FUNCTION_BLOCK IMU_STREAM
  {SET_ATTRIBUTE(OpcUa, SERVICE)}
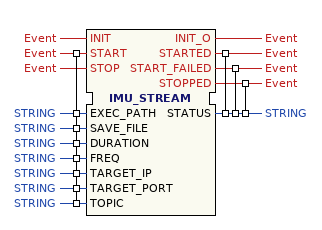
  EVENT_INPUT
    INIT;
    START WITH EXEC_PATH, SAVE_FILE, DURATION, FREQ, TARGET_IP, TARGET_PORT, TOPIC;
    STOP;
  END_EVENT
  EVENT_OUTPUT
    INIT_O;
    STARTED WITH STATUS;
    START_FAILED WITH STATUS;
    STOPPED WITH STATUS;
  END_EVENT
  VAR_INPUT
    EXEC_PATH : STRING; {SET_ATTRIBUTE(OpcUa, Variable)}
    SAVE_FILE : STRING; {SET_ATTRIBUTE(OpcUa, Variable)}
    DURATION : STRING; {SET_ATTRIBUTE(OpcUa, Variable)}
    FREQ : STRING; {SET_ATTRIBUTE(OpcUa, Variable)}
    TARGET_IP : STRING; {SET_ATTRIBUTE(OpcUa, Variable)}
    TARGET_PORT : STRING; {SET_ATTRIBUTE(OpcUa, Variable)}
    TOPIC : STRING; {SET_ATTRIBUTE(OpcUa, Variable)}
  END_VAR
  VAR_OUTPUT
    STATUS : STRING; {SET_ATTRIBUTE(OpcUa, Variable)}
  END_VAR
END_FUNCTION_BLOCK
